// Interpolation strategy used by cmdConvert when building the motion function
// from the raw taught points. Stored raw, so this may change and be regenerated.
TYPE E_CamTeach_Interp :
(
    eLinear  := 0,   // straight segments between points (MOTIONFUNCTYPE_LINEAR)
    eCubicC1 := 1    // POLYNOM3 + central-difference slope -> C1-smooth cubic from position-only teaching
) INT;
END_TYPE

(* stored: Version 1.1.0.1
   DUT E_CamTeach_Interp: Id {0794eda1-2fc4-447f-865e-a5e055910e1c} *)
